// TwinCAT 3 PLC project adc
// ProgramVersion: 3.1.4026.24
// libraries:
//   Tc2_MC2, * (Beckhoff Automation GmbH)
//   Tc2_Standard, * (Beckhoff Automation GmbH)
//   Tc2_System, * (Beckhoff Automation GmbH)
// project tree:
//   DUTs/ E_SlideState.TcDUT
//   GVLs/ GVL_Cfg.TcGVL, GVL_Cmd.TcGVL, GVL_IO.TcGVL, GVL_State.TcGVL
//   / PlcTask.TcTTO
//   POUs/ FB_AdcController.TcPOU, FB_Rotator.TcPOU, FB_RotatorSim.TcPOU, FB_Slide.TcPOU, FB_SlideSim.TcPOU, MAIN.TcPOU
// real-time tasks:
//   TASK PlcTask: cycle T#10ms, priority 20, ADS port 350
//   TASK PlcTask1: cycle T#10ms, priority 21, ADS port 351
// motion (NC):
//   TASK NC-Task 1 SAF: cycle T#2ms, priority 4, ADS port 501
//   TASK NC-Task 1 SVB: cycle T#10ms, priority 8, ADS port 511
//   AXIS Axis 1 (id 1)
//     General: UnitName=°
//     Dynamic: AccelerationMaximum=2000, DecelerationMaximum=2000
//     Velo: Maximum=162
//     OtherSettings: AllowMotionCmdToSlave=true
//     encoder EncType=4
//       EncPara: ScaleFactorNumerator=360, ScaleFactorDenominator=2048, MaxCount=#x0000ffff
//         Inc: RefSyncInverse=false, RefMode=3, RefSoftSyncMask=#x0000ffff
//     drive DrvType=23
//       Analog: VeloReferenz=210, TorqueSetpointScale=10, ScaleFactorActTorque=0.1
//       TimeComp: TaskDelayCycles=1
//     controller CtrType=1
//       CtrPara: PriorControlFactor=1
//         PosDiffControl: Enable=false
//         Observer: BandWidth=20
//   AXIS Axis 2 (id 2)
//     OtherSettings: AllowMotionCmdToSlave=true
//     encoder EncType=4
//       EncPara: MaxCount=#x0000ffff
//         Inc: RefSoftSyncMask=#x0000ffff
//     drive DrvType=23
//       Analog: TorqueSetpointScale=10, ScaleFactorActTorque=0.1
//       TimeComp: TaskDelayCycles=1
//     controller CtrType=1
//       CtrPara: PriorControlFactor=1
//         Observer: BandWidth=20
// I/O:
//   DEVICE Device 1 (EtherCAT), AmsNetId 5.171.247.155.2.1
//     Term 7 (EK1200) [EK1200-5000 EtherCAT Power supply (2A E-Bus)]
//       Term 8 (EL2002) [EL2002 2Ch. Dig. Output 24V, 0.5A]
//       Term 9 (EL1084) [EL1084 4Ch. Dig. Input 24V, 3ms, negative]
//       Term 10 (EL7342) [EL7342 2Ch. DC motor output stage (50V, 3.5A)]
//       Term 11 (EL9505) [EL9505 Power supply terminal 5V]
//       Term 12 (EL9512) [EL9512 Power supply terminal 12V]
//       Term 13 (EL2084) [EL2084 4Ch. Dig. Output 24V, 0.5A, switching to negative]
//       Term 14 (EL9011) [EL9011 End Terminal]
// variable links:
//   adc/adc Instance <-> Device 1 (EtherCAT)/Term 7 (EK1200)/Term 13 (EL2084)
//     PlcTask Outputs/GVL_IO.bMilkyFlat_Out <-> Channel 2/Output
//     PlcTask Outputs/GVL_IO.bShutter_Out <-> Channel 1/Output
//   adc/adc Instance <-> NC-Task 1 SAF/Axes/Axis 1
//     PlcTask Inputs/MAIN.Axis_A_ref.NcToPlc <-> Outputs/ToPlc
//     PlcTask Outputs/MAIN.Axis_A_ref.PlcToNc <-> Inputs/FromPlc
//   adc/adc Instance <-> NC-Task 1 SAF/Axes/Axis 2
//     PlcTask Inputs/MAIN.Axis_B_ref.NcToPlc <-> Outputs/ToPlc
//     PlcTask Outputs/MAIN.Axis_B_ref.PlcToNc <-> Inputs/FromPlc

CONFIGURATION adc
    RESOURCE PLC ON TwinCAT3
        TASK PlcTask(INTERVAL := T#10ms, PRIORITY := 21);
        PROGRAM MAIN WITH PlcTask : MAIN;
    END_RESOURCE
END_CONFIGURATION

// ---- DUTs/E_SlideState.TcDUT
TYPE E_SlideState :
(
    eSlideOut    := 0,
    eSlideIn     := 1,
    eSlideMoving := 2,
    eSlideError  := 3
) INT;
END_TYPE

// ---- GVLs/GVL_Cfg.TcGVL
// Tunables. Persisted in the PLC project, not visible over ADS.
//
// Homing velocity and home position are NOT here — they're NC axis parameters
// set in System Manager (Reference Velocity Fast/Slow, Home Position /
// Calibration Value) at bench bring-up. See docs/bring-up.md § 4.
{attribute 'qualified_only'}
VAR_GLOBAL CONSTANT
    // Default velocity for rotator slews (deg/s). Override per axis if needed.
    rRotatorVelocity  : LREAL := 30.0;
    // Default acceleration / deceleration (deg/s²). Tc2_MC2 takes the same units
    // as the encoder scaling (deg here).
    rRotatorAccel     : LREAL := 60.0;
    rRotatorDecel     : LREAL := 60.0;
    // Jerk (deg/s³). Set to zero to use the NC axis default.
    rRotatorJerk      : LREAL := 0.0;
    // Slide settle timeout — if MOVING persists past this, transition to ERROR.
    tSlideStuckTime   : TIME  := T#5S;
    // Sim-only: how long the simulated slide reports MOVING before settling.
    tSimSlideSettle   : TIME  := T#500MS;
END_VAR

VAR_GLOBAL
    // Sim toggle. TRUE -> FB_AdcController calls FB_*Sim instead of the real FBs.
    // Persist via XAE → "Initialize via retain" or set in the boot project.
    bSimulate : BOOL := FALSE;
END_VAR

// ---- GVLs/GVL_Cmd.TcGVL
// ADS-writable command surface. Python writes here; the PLC consumes and
// clears the edge-triggered bits. The level-triggered slide bits stay set.
{attribute 'qualified_only'}
VAR_GLOBAL

    // Rotator A
    rAxisA_Target : LREAL;
    bAxisA_Go     : BOOL;  // rising edge -> MC_MoveAbsolute; PLC clears after consume
    bAxisA_Stop   : BOOL;  // rising edge -> MC_Stop
    bAxisA_Home   : BOOL;  // rising edge -> MC_Home
    bAxisA_Reset  : BOOL;  // rising edge -> MC_Reset

    // Rotator B
    rAxisB_Target : LREAL;
    bAxisB_Go     : BOOL;
    bAxisB_Stop   : BOOL;
    bAxisB_Home   : BOOL;
    bAxisB_Reset  : BOOL;

    // Slides (level-triggered; TRUE = drive to IN)
    bSlideA_Deploy : BOOL;
    bSlideB_Deploy : BOOL;

    // Shutter & milky-flat diffuser (level-triggered)
    bShutter_Closed   : BOOL;  // TRUE = shutter closed (= EL2084 ch.1 DE-energized)
    bMilkyFlat_Deploy : BOOL;  // TRUE = diffuser in beam (= EL2084 ch.2 DE-energized; wiring is reversed)

END_VAR

// ---- GVLs/GVL_IO.TcGVL
// Hardware-linked I/O. Each variable is bound to an EtherCAT channel via
// TcLinkTo *and* mapped into the process image with AT %I* / AT %Q*.
// If the System Manager topology numbers differ from what's documented
// here, update the path strings (XAE → variable Properties → Path).
//
// Topology (per docs/bring-up.md and bench verification):
//   Term 1 (EK1200) — bus coupler
//   Term 2 (EL2002) — 2-ch DO; ch.1 = Deploy B, ch.2 = Deploy A
//   Term 3 (EL1084) — 4-ch DI; ch.1 = Sense B OUT, ch.2 = Sense B IN,
//                              ch.3 = Sense A OUT, ch.4 = Sense A IN
//   Term 7 (EK1200) — second coupler segment
//   Term 13 (EL2084) — 4-ch DO (negative-switching);
//                              ch.1 = Shutter   (energized = OPEN)
//                              ch.2 = Milky flat (energized = RETRACTED)
//
// Syntax note: the AT %I* (input) or AT %Q* (output) address is REQUIRED
// for TcLinkTo to actually map the variable into the process image. The *
// is a wildcard the compiler resolves at build time. BOOLs link to the
// channel's Input/Output sub-item directly (no '.member :=' prefix).
// Reference:
// https://infosys.beckhoff.com/content/1033/tc3_plc_intro/3107974923.html
{attribute 'qualified_only'}
VAR_GLOBAL

    // --- Slide A: Deploy A on EL2002 ch.2, limits on EL1084 ch.3/4 -----
    {attribute 'TcLinkTo' := 'TIID^Device 1 (EtherCAT)^Term 1 (EK1200)^Term 2 (EL2002)^Channel 2^Output'}
    bSlideA_DeployOut AT %Q* : BOOL;

    {attribute 'TcLinkTo' := 'TIID^Device 1 (EtherCAT)^Term 1 (EK1200)^Term 3 (EL1084)^Channel 4^Input'}
    bSlideA_LimitIn AT %I* : BOOL;

    {attribute 'TcLinkTo' := 'TIID^Device 1 (EtherCAT)^Term 1 (EK1200)^Term 3 (EL1084)^Channel 3^Input'}
    bSlideA_LimitOut AT %I* : BOOL;

    // --- Slide B: Deploy B on EL2002 ch.1, limits on EL1084 ch.1/2 -----
    {attribute 'TcLinkTo' := 'TIID^Device 1 (EtherCAT)^Term 1 (EK1200)^Term 2 (EL2002)^Channel 1^Output'}
    bSlideB_DeployOut AT %Q* : BOOL;

    {attribute 'TcLinkTo' := 'TIID^Device 1 (EtherCAT)^Term 1 (EK1200)^Term 3 (EL1084)^Channel 2^Input'}
    bSlideB_LimitIn AT %I* : BOOL;

    {attribute 'TcLinkTo' := 'TIID^Device 1 (EtherCAT)^Term 1 (EK1200)^Term 3 (EL1084)^Channel 1^Input'}
    bSlideB_LimitOut AT %I* : BOOL;

    // --- Shutter & milky-flat diffuser: EL2084 on the second coupler ----
    // EL2084 is the NEGATIVE-switching 4-ch DO variant (switches 0 V, not
    // +24 V) — verify actuator wiring/polarity on the bench before relying
    // on TRUE = energized.
    {attribute 'TcLinkTo' := 'TIID^Device 1 (EtherCAT)^Term 7 (EK1200)^Term 13 (EL2084)^Channel 1^Output'}
    bShutter_Out AT %Q* : BOOL;

    {attribute 'TcLinkTo' := 'TIID^Device 1 (EtherCAT)^Term 7 (EK1200)^Term 13 (EL2084)^Channel 2^Output'}
    bMilkyFlat_Out AT %Q* : BOOL;

    // Rotator axes (EL7342 channels) are bound via the NC axis configuration,
    // not via GVL_IO. See docs/bring-up.md § 3.

END_VAR

// ---- GVLs/GVL_State.TcGVL
// ADS-readable telemetry. Mirrors plc_client.py _AXIS_SYMBOLS / _SLIDE_SYMBOLS.
// Treat as read-only from the Python side.
{attribute 'qualified_only'}
VAR_GLOBAL

    // Rotator A
    rAxisA_Position : LREAL;
    bAxisA_Busy     : BOOL;
    bAxisA_Done     : BOOL;
    bAxisA_Error    : BOOL;
    nAxisA_ErrorId  : UDINT;  // Matches MC_*.ErrorID (Tc2_MC2)
    bAxisA_Ready    : BOOL;   // Homed AND not in error — see FB_Rotator.bReady

    // Rotator B
    rAxisB_Position : LREAL;
    bAxisB_Busy     : BOOL;
    bAxisB_Done     : BOOL;
    bAxisB_Error    : BOOL;
    nAxisB_ErrorId  : UDINT;
    bAxisB_Ready    : BOOL;

    // Slides
    eSlideA : E_SlideState;
    eSlideB : E_SlideState;

    // Shutter & milky-flat diffuser. No position feedback on either — these
    // echo the commanded state, not a measured one.
    bShutter_Closed     : BOOL;
    bMilkyFlat_Deployed : BOOL;

    // Heartbeat: toggled every cycle by MAIN. Python uses it for liveness.
    bHeartbeat : BOOL;

END_VAR

// ---- POUs/MAIN.TcPOU
// PLC entry point. Single FB_AdcController instance does all the work.
//
// Axis_A_ref / Axis_B_ref are linked to the NC axes via the System Manager:
// MOTION → NC-Task → Axis A/B → right-click → "Change Link" → bind to these
// AXIS_REF instances. See docs/bring-up.md § 3.

PROGRAM MAIN
VAR
    fbAdc : FB_AdcController;

    // Link these to the NC axes in System Manager.
    Axis_A_ref : AXIS_REF;
    Axis_B_ref : AXIS_REF;

    // Task cycle in seconds. Keep in sync with the task period configured
    // in XAE (default 10ms here).
    rCycleSeconds : LREAL := 0.010;
END_VAR

fbAdc(
    AxisA := Axis_A_ref,
    AxisB := Axis_B_ref,
    rCycleSeconds := rCycleSeconds
);

END_PROGRAM

// ---- POUs/FB_AdcController.TcPOU
// Composition root. Owns both rotator instances (real + sim) and both slide
// instances (real + sim) per axis. Each cycle, dispatches to the appropriate
// variant based on GVL_Cfg.bSimulate.
//
// All GVL_State / GVL_Cmd reads and writes happen here — no other POU should
// touch them. This keeps the ADS-visible state machine concentrated in one
// place.
//
// The real rotators take AXIS_REFs from the NC config. Wire them in MAIN.

FUNCTION_BLOCK FB_AdcController
VAR_IN_OUT
    AxisA : AXIS_REF;
    AxisB : AXIS_REF;
END_VAR
VAR_INPUT
    rCycleSeconds : LREAL;
END_VAR
VAR
    fbRotatorA     : FB_Rotator;
    fbRotatorB     : FB_Rotator;
    fbRotatorSimA  : FB_RotatorSim;
    fbRotatorSimB  : FB_RotatorSim;
    fbSlideA       : FB_Slide;
    fbSlideB       : FB_Slide;
    fbSlideSimA    : FB_SlideSim;
    fbSlideSimB    : FB_SlideSim;
END_VAR

// --- Rotator A ---------------------------------------------------------
IF GVL_Cfg.bSimulate THEN
    fbRotatorSimA(
        bGo := GVL_Cmd.bAxisA_Go,
        rTarget := GVL_Cmd.rAxisA_Target,
        rVelocity := GVL_Cfg.rRotatorVelocity,
        bStop := GVL_Cmd.bAxisA_Stop,
        bHome := GVL_Cmd.bAxisA_Home,
        bReset := GVL_Cmd.bAxisA_Reset,
        rCycleSeconds := rCycleSeconds
    );
    GVL_State.rAxisA_Position := fbRotatorSimA.rPosition;
    GVL_State.bAxisA_Busy     := fbRotatorSimA.bBusy;
    GVL_State.bAxisA_Done     := fbRotatorSimA.bDone;
    GVL_State.bAxisA_Error    := fbRotatorSimA.bError;
    GVL_State.nAxisA_ErrorId  := fbRotatorSimA.nErrorId;
    GVL_State.bAxisA_Ready    := fbRotatorSimA.bReady;
ELSE
    fbRotatorA(
        Axis := AxisA,
        bGo := GVL_Cmd.bAxisA_Go,
        rTarget := GVL_Cmd.rAxisA_Target,
        rVelocity := GVL_Cfg.rRotatorVelocity,
        rAccel := GVL_Cfg.rRotatorAccel,
        rDecel := GVL_Cfg.rRotatorDecel,
        rJerk := GVL_Cfg.rRotatorJerk,
        bStop := GVL_Cmd.bAxisA_Stop,
        bHome := GVL_Cmd.bAxisA_Home,
        bReset := GVL_Cmd.bAxisA_Reset
    );
    GVL_State.rAxisA_Position := fbRotatorA.rPosition;
    GVL_State.bAxisA_Busy     := fbRotatorA.bBusy;
    GVL_State.bAxisA_Done     := fbRotatorA.bDone;
    GVL_State.bAxisA_Error    := fbRotatorA.bError;
    GVL_State.nAxisA_ErrorId  := fbRotatorA.nErrorId;
    GVL_State.bAxisA_Ready    := fbRotatorA.bReady;
END_IF

// The PLC clears the Go bit after one cycle so the next rising edge can fire.
GVL_Cmd.bAxisA_Go    := FALSE;
GVL_Cmd.bAxisA_Stop  := FALSE;
GVL_Cmd.bAxisA_Home  := FALSE;
GVL_Cmd.bAxisA_Reset := FALSE;

// --- Rotator B ---------------------------------------------------------
IF GVL_Cfg.bSimulate THEN
    fbRotatorSimB(
        bGo := GVL_Cmd.bAxisB_Go,
        rTarget := GVL_Cmd.rAxisB_Target,
        rVelocity := GVL_Cfg.rRotatorVelocity,
        bStop := GVL_Cmd.bAxisB_Stop,
        bHome := GVL_Cmd.bAxisB_Home,
        bReset := GVL_Cmd.bAxisB_Reset,
        rCycleSeconds := rCycleSeconds
    );
    GVL_State.rAxisB_Position := fbRotatorSimB.rPosition;
    GVL_State.bAxisB_Busy     := fbRotatorSimB.bBusy;
    GVL_State.bAxisB_Done     := fbRotatorSimB.bDone;
    GVL_State.bAxisB_Error    := fbRotatorSimB.bError;
    GVL_State.nAxisB_ErrorId  := fbRotatorSimB.nErrorId;
    GVL_State.bAxisB_Ready    := fbRotatorSimB.bReady;
ELSE
    fbRotatorB(
        Axis := AxisB,
        bGo := GVL_Cmd.bAxisB_Go,
        rTarget := GVL_Cmd.rAxisB_Target,
        rVelocity := GVL_Cfg.rRotatorVelocity,
        rAccel := GVL_Cfg.rRotatorAccel,
        rDecel := GVL_Cfg.rRotatorDecel,
        rJerk := GVL_Cfg.rRotatorJerk,
        bStop := GVL_Cmd.bAxisB_Stop,
        bHome := GVL_Cmd.bAxisB_Home,
        bReset := GVL_Cmd.bAxisB_Reset
    );
    GVL_State.rAxisB_Position := fbRotatorB.rPosition;
    GVL_State.bAxisB_Busy     := fbRotatorB.bBusy;
    GVL_State.bAxisB_Done     := fbRotatorB.bDone;
    GVL_State.bAxisB_Error    := fbRotatorB.bError;
    GVL_State.nAxisB_ErrorId  := fbRotatorB.nErrorId;
    GVL_State.bAxisB_Ready    := fbRotatorB.bReady;
END_IF

GVL_Cmd.bAxisB_Go    := FALSE;
GVL_Cmd.bAxisB_Stop  := FALSE;
GVL_Cmd.bAxisB_Home  := FALSE;
GVL_Cmd.bAxisB_Reset := FALSE;

// --- Slide A ----------------------------------------------------------
IF GVL_Cfg.bSimulate THEN
    fbSlideSimA(bDeploy := GVL_Cmd.bSlideA_Deploy, tSettle := GVL_Cfg.tSimSlideSettle);
    GVL_State.eSlideA := fbSlideSimA.eState;
    GVL_IO.bSlideA_DeployOut := FALSE;  // never assert real output in sim
ELSE
    fbSlideA(
        bDeploy := GVL_Cmd.bSlideA_Deploy,
        bLimitIn := GVL_IO.bSlideA_LimitIn,
        bLimitOut := GVL_IO.bSlideA_LimitOut,
        tStuck := GVL_Cfg.tSlideStuckTime
    );
    GVL_State.eSlideA := fbSlideA.eState;
    GVL_IO.bSlideA_DeployOut := fbSlideA.bSolenoid;
END_IF

// --- Slide B ----------------------------------------------------------
IF GVL_Cfg.bSimulate THEN
    fbSlideSimB(bDeploy := GVL_Cmd.bSlideB_Deploy, tSettle := GVL_Cfg.tSimSlideSettle);
    GVL_State.eSlideB := fbSlideSimB.eState;
    GVL_IO.bSlideB_DeployOut := FALSE;
ELSE
    fbSlideB(
        bDeploy := GVL_Cmd.bSlideB_Deploy,
        bLimitIn := GVL_IO.bSlideB_LimitIn,
        bLimitOut := GVL_IO.bSlideB_LimitOut,
        tStuck := GVL_Cfg.tSlideStuckTime
    );
    GVL_State.eSlideB := fbSlideB.eState;
    GVL_IO.bSlideB_DeployOut := fbSlideB.bSolenoid;
END_IF

// --- Shutter ----------------------------------------------------------
// Plain DO, no position feedback. Energizing EL2084 ch.1 OPENS the
// shutter, so bShutter_Closed = TRUE drives the output FALSE. State
// echoes the command; in sim the real output stays de-energized (same
// convention as the slides).
IF GVL_Cfg.bSimulate THEN
    GVL_IO.bShutter_Out := FALSE;
ELSE
    GVL_IO.bShutter_Out := NOT GVL_Cmd.bShutter_Closed;
END_IF
GVL_State.bShutter_Closed := GVL_Cmd.bShutter_Closed;

// --- Milky-flat diffuser ----------------------------------------------
// Reversed wiring: energizing EL2084 ch.2 RETRACTS the diffuser, so
// deploy = output de-energized. In sim the real output still stays FALSE.
IF GVL_Cfg.bSimulate THEN
    GVL_IO.bMilkyFlat_Out := FALSE;
ELSE
    GVL_IO.bMilkyFlat_Out := NOT GVL_Cmd.bMilkyFlat_Deploy;
END_IF
GVL_State.bMilkyFlat_Deployed := GVL_Cmd.bMilkyFlat_Deploy;

// Heartbeat — flipped here so Python sees it tick every cycle.
GVL_State.bHeartbeat := NOT GVL_State.bHeartbeat;

END_FUNCTION_BLOCK

// ---- POUs/FB_Rotator.TcPOU
// Real rotator. Wraps Tc2_MC2 against an NC axis. The Go/Stop/Home/Reset
// inputs are edge-triggered to mirror the ADS command semantics.
//
// Homing uses MC_Home with bCalibrationCam driven from the PLC — Beckhoff's
// documented pattern for axes with only an encoder sync pulse (no physical
// reference cam). NC's two-phase homing model is preserved; the PLC simulates
// a permanently-occupied cam during Phase 1 (search), and NC's configured
// Reference Mode (e.g. Hardware Latch 1) captures the precise position in
// Phase 2 via the EL7342 external latch on I1 / I2.
//
// Reference: Tc2_MC2 MC_Home documentation —
//   https://infosys.beckhoff.com/content/1033/tcplclib_tc2_mc2/70117515.html
//   "If an axis is to be referenced without referencing cam, i.e. only based
//    on the sync pulse of the encoder, the referencing cam can be simulated
//    via the PLC program. The 'bCalibrationCam' signal is initially activated
//    and then canceled, if Axis.NcToPlc.HomingState is equal or greater 4."
//
// NC bench-time configuration (System Manager → NC → Axis → Encoder):
//   Reference Mode (Sync condition) = Hardware Latch 1 (pos. edge)
//   Invert Direction for Sync Impulse Search = FALSE  (Z is active-high on I1)
//   Reference Velocity (Fast) / (Slow) — bench-tuned values
//   Home Position (Calibration Value) — final position written after sync

FUNCTION_BLOCK FB_Rotator
VAR_IN_OUT
    Axis : AXIS_REF;
END_VAR
VAR_INPUT
    bGo       : BOOL;
    rTarget   : LREAL;
    rVelocity : LREAL;
    rAccel    : LREAL;
    rDecel    : LREAL;
    rJerk     : LREAL;
    bStop     : BOOL;
    bHome     : BOOL;
    bReset    : BOOL;
END_VAR
VAR_OUTPUT
    rPosition : LREAL;
    bBusy     : BOOL;
    bDone     : BOOL;
    bError    : BOOL;
    nErrorId  : UDINT;
    // Ready = axis has been homed at least once since boot AND is not in error.
    // The intended use is gating: any caller that needs absolute position
    // should refuse to dispatch a move when bReady = FALSE.
    bReady    : BOOL;
END_VAR
VAR
    fbPower    : MC_Power;
    fbMove     : MC_MoveAbsolute;
    fbStop     : MC_Stop;
    fbHome     : MC_Home;
    fbReset    : MC_Reset;
    fbReadPos  : MC_ReadActualPosition;
    fbStatus   : MC_ReadStatus;
    rfGo       : R_TRIG;
    rfStop     : R_TRIG;
    rfHome     : R_TRIG;
    rfReset    : R_TRIG;
    bHomed     : BOOL;     // latched TRUE once a homing run completes successfully
END_VAR

// Always enabled. Override per-axis safety in the NC config, not here.
fbPower(
    Axis            := Axis,
    Enable          := TRUE,
    Enable_Positive := TRUE,
    Enable_Negative := TRUE,
    Override        := 100.0
);

// Edge detection on the commands.
rfGo(CLK := bGo);
rfStop(CLK := bStop);
rfHome(CLK := bHome);
rfReset(CLK := bReset);

// Reset clears latched errors first so the next Go can run.
fbReset(Axis := Axis, Execute := rfReset.Q);

// Stop aborts everything, including a running homing sequence.
fbStop(Axis := Axis, Execute := rfStop.Q, Deceleration := rDecel);

// Homing — Beckhoff's documented cam-less pattern for axes with only an
// encoder Z (no physical reference cam): drive MC_Home.bCalibrationCam from
// the PLC to simulate a permanently-occupied cam through Phase 1, then let
// NC's configured Reference Mode (Hardware Latch 1, pos. edge for the
// active-high Z directly on I1) capture the precise position in Phase 2.
fbHome(
    Axis            := Axis,
    Execute         := rfHome.Q,
    Position        := 0.0,
    HomingMode      := MC_DefaultHoming,
    BufferMode      := MC_Aborting,
    bCalibrationCam :=  Axis.NcToPlc.HomingState < 4
);

fbMove(
    Axis         := Axis,
    Execute      := rfGo.Q,
    Position     := rTarget,
    Velocity     := rVelocity,
    Acceleration := rAccel,
    Deceleration := rDecel,
    Jerk         := rJerk,
    BufferMode   := MC_Aborting
);

// Live readback.
fbReadPos(Axis := Axis, Enable := TRUE);
fbStatus(Axis := Axis, Enable := TRUE);

rPosition := fbReadPos.Position;
// MC_ReadStatus has no .Moving flag; the action-FB Busy bits cover all motion.
bBusy     := fbMove.Busy OR fbHome.Busy OR fbStop.Busy;
bDone     := (fbMove.Done OR fbHome.Done) AND NOT bBusy;

// Latch bHomed. NC clears HomingState back to 0 once MC_Home finishes, so we
// can't infer "homed" from HomingState directly. Instead we set the latch on
// fbHome.Done and clear it on the next rfHome rising edge (axis is no longer
// calibrated while a new homing run is in progress). A reset doesn't clear
// bHomed — the mechanical calibration survives an error/reset cycle.
IF rfHome.Q THEN
    bHomed := FALSE;
END_IF
IF fbHome.Done AND NOT fbHome.Error THEN
    bHomed := TRUE;
END_IF

bReady := bHomed AND NOT bError;

// Bubble up the first error we find.
IF fbMove.Error THEN
    bError := TRUE; nErrorId := fbMove.ErrorID;
ELSIF fbHome.Error THEN
    bError := TRUE; nErrorId := fbHome.ErrorID;
ELSIF fbStop.Error THEN
    bError := TRUE; nErrorId := fbStop.ErrorID;
ELSIF fbReset.Error THEN
    bError := TRUE; nErrorId := fbReset.ErrorID;
ELSIF fbPower.Error THEN
    bError := TRUE; nErrorId := fbPower.ErrorID;
ELSE
    bError := FALSE; nErrorId := 0;
END_IF

END_FUNCTION_BLOCK

// ---- POUs/FB_RotatorSim.TcPOU
// Software-only rotator. Same interface as FB_Rotator (minus the AXIS_REF),
// integrates position toward target at rVelocity. No real motion is asserted.
FUNCTION_BLOCK FB_RotatorSim
VAR_INPUT
    bGo           : BOOL;
    rTarget       : LREAL;
    rVelocity     : LREAL;
    bStop         : BOOL;
    bHome         : BOOL;
    bReset        : BOOL;
    rCycleSeconds : LREAL;   // task cycle in seconds (e.g. 0.010)
END_VAR
VAR_OUTPUT
    rPosition : LREAL;
    bBusy     : BOOL;
    bDone     : BOOL;
    bError    : BOOL;
    nErrorId  : UDINT;
    bReady    : BOOL;       // homed AND not in error (sim mirrors FB_Rotator)
END_VAR
VAR
    rActiveTarget : LREAL;
    rDelta        : LREAL;
    rMaxStep      : LREAL;
    rfGo          : R_TRIG;
    rfStop        : R_TRIG;
    rfHome        : R_TRIG;
    rfReset       : R_TRIG;
    bSimHomed     : BOOL := FALSE;   // latched on first bHome rising edge
END_VAR

rfGo(CLK := bGo);
rfStop(CLK := bStop);
rfHome(CLK := bHome);
rfReset(CLK := bReset);

IF rfReset.Q THEN
    bError := FALSE;
    nErrorId := 0;
END_IF

IF rfHome.Q THEN
    // Home is the absolute zero in sim. The real axis uses the NC Reference
    // Position parameter set in System Manager — bench-time configuration.
    rPosition := 0.0;
    rActiveTarget := 0.0;
    bBusy := FALSE;
    bDone := TRUE;
    bSimHomed := TRUE;
END_IF

bReady := bSimHomed AND NOT bError;

IF rfStop.Q THEN
    rActiveTarget := rPosition;
    bBusy := FALSE;
    bDone := TRUE;
END_IF

IF rfGo.Q THEN
    rActiveTarget := rTarget;
    bBusy := TRUE;
    bDone := FALSE;
END_IF

// Advance toward the active target at rVelocity * dt per cycle.
IF bBusy THEN
    rDelta := rActiveTarget - rPosition;
    rMaxStep := rVelocity * rCycleSeconds;
    IF ABS(rDelta) <= rMaxStep THEN
        rPosition := rActiveTarget;
        bBusy := FALSE;
        bDone := TRUE;
    ELSIF rDelta > 0.0 THEN
        rPosition := rPosition + rMaxStep;
    ELSE
        rPosition := rPosition - rMaxStep;
    END_IF
END_IF

END_FUNCTION_BLOCK

// ---- POUs/FB_Slide.TcPOU
// Real pneumatic slide. Drives the solenoid output when bDeploy=TRUE,
// reports state via limit switches with a stuck-detection timer.
FUNCTION_BLOCK FB_Slide
VAR_INPUT
    bDeploy   : BOOL;        // level: TRUE = drive to IN
    bLimitIn  : BOOL;
    bLimitOut : BOOL;
    tStuck    : TIME;        // moving longer than this -> ERROR
END_VAR
VAR_OUTPUT
    bSolenoid : BOOL;        // drives the EL2002 channel
    eState    : E_SlideState;
END_VAR
VAR
    tonStuck : TON;
END_VAR

// Solenoid drive is a direct mirror of the deploy request.
bSolenoid := bDeploy;

// Decode state from limit switches.
IF bLimitIn AND NOT bLimitOut THEN
    eState := E_SlideState.eSlideIn;
    tonStuck(IN := FALSE);
ELSIF bLimitOut AND NOT bLimitIn THEN
    eState := E_SlideState.eSlideOut;
    tonStuck(IN := FALSE);
ELSIF bLimitIn AND bLimitOut THEN
    // Both switches asserted simultaneously -> wiring fault.
    eState := E_SlideState.eSlideError;
    tonStuck(IN := FALSE);
ELSE
    // Neither switch asserted -> mid-travel.
    eState := E_SlideState.eSlideMoving;
    tonStuck(IN := TRUE, PT := tStuck);
    IF tonStuck.Q THEN
        eState := E_SlideState.eSlideError;
    END_IF
END_IF

END_FUNCTION_BLOCK

// ---- POUs/FB_SlideSim.TcPOU
// Software-only slide. Same outputs as FB_Slide; ignores hardware inputs.
// Transitions through MOVING for tSettle ms after bDeploy changes.
FUNCTION_BLOCK FB_SlideSim
VAR_INPUT
    bDeploy : BOOL;
    tSettle : TIME;
END_VAR
VAR_OUTPUT
    bSolenoid : BOOL;       // not wired; provided for interface parity
    eState    : E_SlideState;
END_VAR
VAR
    bDeployPrev : BOOL;
    bSettling   : BOOL;
    bTargetIn   : BOOL;
    tonSettle   : TON;
END_VAR

bSolenoid := bDeploy;

// Detect a change in the requested position.
IF bDeploy <> bDeployPrev THEN
    bDeployPrev := bDeploy;
    bTargetIn := bDeploy;
    bSettling := TRUE;
    tonSettle(IN := FALSE);
END_IF

IF bSettling THEN
    tonSettle(IN := TRUE, PT := tSettle);
    eState := E_SlideState.eSlideMoving;
    IF tonSettle.Q THEN
        bSettling := FALSE;
        tonSettle(IN := FALSE);
    END_IF
ELSE
    IF bTargetIn THEN
        eState := E_SlideState.eSlideIn;
    ELSE
        eState := E_SlideState.eSlideOut;
    END_IF
END_IF

END_FUNCTION_BLOCK
